# EPICS autosave request: 1.5.0/debian-12/7.0.10/modules/ADCore-ee039d2/db/NDPluginBase_settings.req
$(P)$(R)NDArrayPort
$(P)$(R)NDArrayAddress
$(P)$(R)EnableCallbacks
$(P)$(R)MinCallbackTime
$(P)$(R)MaxByteRate
$(P)$(R)BlockingCallbacks
$(P)$(R)QueueSize
$(P)$(R)NumThreads
$(P)$(R)SortTime
$(P)$(R)SortMode
$(P)$(R)SortSize
file "NDArrayBase_settings.req", P=$(P), R=$(R)
